Fanuc KAREL source: kc00042.KL

-- PROVISIONAL review KL for V1013-1; original PC SHA256 ebcebea82c46e15118e166269727083992b7dddfca9d8205e14658caa7c6fa2d
-- Incomplete behavior may be omitted. Consult companion uncertainty JSON. Do not deploy.
PROGRAM KC00042
%NOLOCKGROUP
BEGIN
  -- UNRESOLVED_PC offsets 5-35; opcodes 27,22,22,27,9D,31,7E,4A
  -- UNRESOLVED_PC offsets 40-44; opcodes 7F
END KC00042
